ADAPTER LinkSafeSequenceSequenceServices
  (* Standard: 61499-2 *)
  (* Version 3.0, 2026-11-12, sorting2n, sorting2n *)
  PACKAGE Main;
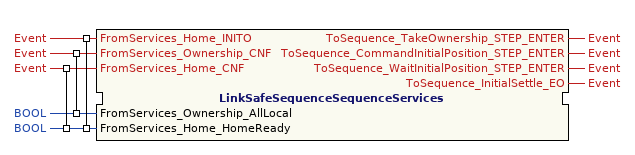
  EVENT_INPUT
    FromServices_Home_INITO WITH FromServices_Home_HomeReady;
    FromServices_Ownership_CNF WITH FromServices_Ownership_AllLocal;
    FromServices_Home_CNF WITH FromServices_Home_HomeReady;
  END_EVENT
  EVENT_OUTPUT
    ToSequence_TakeOwnership_STEP_ENTER;
    ToSequence_CommandInitialPosition_STEP_ENTER;
    ToSequence_WaitInitialPosition_STEP_ENTER;
    ToSequence_InitialSettle_EO;
  END_EVENT
  VAR_INPUT
    FromServices_Ownership_AllLocal : BOOL;
    FromServices_Home_HomeReady : BOOL;
  END_VAR
END_ADAPTER
